{attribute 'qualified_only'}
{attribute 'strict'}
TYPE E_CIP_Mode :
(
	eOff :=0,
	eManual,
	eAuto	
);
END_TYPE

(* stored: Version 1.1.0.1, ProductVersion 3.1.4024.12
   DUT E_CIP_Mode: Id {d8d99f73-1280-477f-982f-8d0ca4e555a3} *)
